{attribute 'qualified_only'}
{attribute 'strict'}
TYPE E_Piston_Recipe_State :
(
	NoChanges := 0,
	Act,	// action invert deafult cmd
	Release	// action deafult cmd
);
END_TYPE

(* stored: Version 1.1.0.1, ProductVersion 3.1.4024.12
   DUT E_Piston_Recipe_State: Id {1f711998-f58d-4a3c-be0c-55264542a250} *)
